(* IEC 61131-3 sources: rungstone/fixtures/plc/two_tank/openplc, 1 file *)

(* ---- two_tank_openplc.st ---- *)
(* GENERATED BY Rungstone - DRAFT FOR ENGINEER REVIEW - NOT APPROVED.
   Test translation of fixtures/plc/two_tank/two_tank_slc.txt (SLC 5/04 ladder file 2) for OpenPLC Runtime.
   Upload through the OpenPLC Runtime Programs page; not for use on a production system without review and testing. *)

PROGRAM prog_TwoTank
  VAR
    Start_PB AT %IX0.0 : BOOL;     (* was I:1/14 start pushbutton (NO) *)
    Stop_PB AT %IX0.1 : BOOL;      (* was I:1/15 stop pushbutton, normally closed: TRUE = not pressed *)
    Tank1_LLS AT %IX0.2 : BOOL;    (* was I:1/0 tank 1 low level switch (TRUE = liquid present) INFERRED *)
    Tank2_LLS AT %IX0.3 : BOOL;    (* was I:1/1 tank 2 low level switch INFERRED *)
    Level_Raw AT %IW0 : UINT;      (* was I:3.0 level transmitter raw; OpenPLC analog input 0..65535 (board-specific) *)
    Master_Run AT %QX0.0 : BOOL;   (* was O:2/15 master coil *)
    Valve1_AO AT %QW0 : UINT;      (* was O:4.0 tank 1 drain valve analog output *)
    Valve2_AO AT %QW1 : UINT;      (* was O:6.0 tank 2 drain valve analog output *)
    Level_Cutoff AT %MW0 : INT;    (* was N7:1 drain cutoff 0..1000, written by the HMI over Modbus (holding register 1024) *)
    Drain_Cmd AT %MW1 : UINT;      (* was N7:2 drain valve command, written by the HMI (holding register 1025) *)
  END_VAR
  VAR
    Level_Pct : INT;               (* was N7:0 scaled level 0..1000 *)
  END_VAR

  (* rung 0: master start/stop seal-in *)
  Master_Run := (Start_PB OR Master_Run) AND Stop_PB;
  (* rung 1: scale level 0..65535 -> 0..1000 *)
  IF Master_Run THEN
    Level_Pct := REAL_TO_INT(UINT_TO_REAL(Level_Raw) * 1000.0 / 65535.0);
  END_IF;
  (* rungs 2-3: drain tank 1 *)
  IF Master_Run AND Tank1_LLS AND Level_Pct > Level_Cutoff THEN
    Valve1_AO := Drain_Cmd;
  END_IF;
  IF NOT Master_Run OR NOT Tank1_LLS OR Level_Pct <= Level_Cutoff THEN
    Valve1_AO := 0;
  END_IF;
  (* rungs 4-5: then drain tank 2 *)
  IF Master_Run AND NOT Tank1_LLS AND Tank2_LLS THEN
    Valve2_AO := Drain_Cmd;
  END_IF;
  IF NOT Master_Run OR NOT Tank2_LLS OR Tank1_LLS THEN
    Valve2_AO := 0;
  END_IF;
END_PROGRAM

CONFIGURATION Config0
  RESOURCE Res0 ON PLC
    TASK Main(INTERVAL := T#10ms, PRIORITY := 0);
    PROGRAM Inst0 WITH Main : prog_TwoTank;
  END_RESOURCE
END_CONFIGURATION
